Staubli VAL3: utCommon.dtx

public string sSourceImage
public string sID
public string sClass
public string sPage
